(* IEC 61131-3 sources: HappyLearnCodesys/content/softmotion/CNC04_table, 2 files *)

(* ---- Ipo.st ---- *)
PROGRAM Ipo
VAR
	trafo: SMC_TRAFO_Gantry2;
	p1,p2: SMC_ControlAxisByPos;
	trafof: SMC_TRAFOF_Gantry2;
	smci: SMC_Interpolator;
	mcp1, mcp2: MC_Power;
END_VAR

(* ---- Path.st ---- *)
PROGRAM Path
VAR
	dec: SMC_NCDecoder;
	SmoothPath: SMC_SmoothPath;
	CheckVel: SMC_CheckVelocities;
	buf1: ARRAY[0..15] OF SMC_GEOINFO;
	buf2: ARRAY[0..99] OF SMC_GEOINFO;
END_VAR
